Fanuc KAREL source: KT00232.KL

PROGRAM KT00232
%NOLOCKGROUP
VAR
  B1: BOOLEAN
  H2: ARRAY[2] OF SHORT
  OUT: INTEGER
BEGIN
  B1 = TRUE
    H2[1] = 3
  OUT = B1 OR H2[1]
END KT00232
